TYPE ST_YASKAWA_REF_1 : FB_YASKAWA_REF;
END_TYPE

(* stored: Version 1.1.0.1, ProductVersion 3.1.4024.15
   DUT ST_YASKAWA_REF_1: Id {75dca1bd-78d0-491c-9dc4-a1ee03cc5249} *)
